// TIA Portal V21 export
// export: Created 2026-11-10T07:02:25.9271257Z, ExportSetting WithDefaults, DisplayName Totally Integrated Automation Portal, DisplayVersion V21 Update 3, DisplayName STEP 7 Professional, DisplayVersion V21 Update 3, DisplayName STEP 7 Safety, DisplayVersion V21, DisplayName Tech WebApplication, DisplayVersion V21, DisplayName WinCC Basic/Comfort/Advanced, DisplayVersion V21 Update 3, DisplayName WinCC Unified, DisplayVersion V21 Update 3
FUNCTION "FC_SclStr" : Void   // FC8, SCL
{ S7_Optimized_Access := 'TRUE' }
VERSION : 0.1
// stored: AutoNumber true, IsIECCheckEnabled false, SetENOAutomatically false, UDAEnableTagReadback false
   VAR_TEMP
      s : String;
      s2 : String;
      ws : WString;
      i : Int;
      c : Char;
      "b" : Bool;
      r : Real;
   END_VAR
BEGIN
   #i := LEN(#s);
   #s := CONCAT(IN1 := #s, IN2 := #s2);
   #s := LEFT(IN := #s, L := 2);
   #s := RIGHT(IN := #s, L := 2);
   #s := MID(IN := #s, L := 2, P := 1);
   #i := FIND(IN1 := #s, IN2 := #s2);
   #s := INSERT(IN1 := #s, IN2 := #s2, P := 1);
   #s := DELETE(IN := #s, L := 1, P := 1);
   #s := REPLACE(IN1 := #s, IN2 := #s2, L := 1, P := 1);
   #b := #s = #s2;
   #b := #s <> #s2;
   #b := #s < #s2;
   #c := #s[1];
   #s[1] := #c;
   #s := INT_TO_STRING(#i);
   #i := STRING_TO_INT(#s);
   #s := REAL_TO_STRING(#r);
   #ws := STRING_TO_WSTRING(#s);
END_FUNCTION
